// TIA Portal project "项目8" (V15.1)

(* hardware
DEVICE "GSD device_1"  GSD.Device.PN
   slot 0: "机架"  Rack  V1.0
   slot 0: "SINAMICS-G120SV-PN"  SINAMICS G120 CU250S-2 PN Vector V4.7  6SL3 246-0BA22-1FAx  V4.70
      slot 0: "SINAMICS G120 CU250S-2 PN Vector V4.7"  SINAMICS G120 CU250S-2 PN Vector V4.7
      slot 1: "DO 矢量_1"  DO VECTOR
         slot 0: "模块访问点"  Module Access Point
      slot 1: "PN-IO"  PN-IO
         slot 1: "端口1"  Port 1
         slot 2: "端口2"  Port 2
   slot 2: "标准报文1, PZD-2/2"  Standard telegram 1, PZD-2/2
DEVICE "S7-1200 station_1"  S7-1200 Station
   slot 0: "Rack_0"  S7-1200 Rack  Rack  V1.0
   slot 1: "PLC_1"  CPU 1214C DC/DC/DC  6ES7 214-1AG40-0XB0  V4.2
   slot 2: "DI 16/DQ 16x24VDC_1"  6ES7 223-1BL32-0XB0  V2.0
   slot 3: "AI 4x13BIT/AQ 2x14BIT_1"  6ES7 234-4HE32-0XB0  V2.0
DEVICE "HMI_1"  KTP700 Basic PN
   slot 0: "HMI_1"  KTP700 Basic PN  6AV2 123-2GB03-0AX0  15.1.0.0
   slot 1: "HMI_RT_1"  KTP700 Basic PN  6AV2 123-2GB03-0AX0  15.1.0.0
   slot 5: "HMI_1.IE_CP_1"  PROFINET Interface  15.0.1.0
      slot 1: "PROFINET Interface_1"  PROFINET Interface
         slot 1: "Port_1"  Port
*)

// ===== PLC "PLC_1"  CPU 1214C DC/DC/DC =====

VAR_GLOBAL   // PLC tag table "默认变量表"
   "G120输出速度" AT %MW0 : Word;
   "G120控制" AT %QW64 : Word;
   "Tag_5" AT %MW12 : Word;
   "G120速度" AT %QW66 : Word;
   "停止" AT %I0.1 : Bool;
   "正转" AT %I0.2 : Bool;
   "反转" AT %I0.3 : Bool;
   "轴_1_脉冲" AT %Q0.0 : Bool;
   "轴_1_方向" AT %Q0.1 : Bool;
   "开关4" AT %I0.4 : Bool;
   "步进电机启动" AT %Q1.0 : Bool;
   "速度" AT %MD10 : Real;
   "32位速度" AT %MD14 : DInt;
   "16位速度" AT %MW18 : UInt;
   "计算速度" AT %MD20 : Real;
   "sds" AT %MW24 : Int;
END_VAR

DATA_BLOCK "轴_1"   // DB1, Motion_DB
{ S7_Optimized_Access := 'TRUE' }
AUTHOR : SIMATIC
FAMILY : BasicMC
NAME : TO_PosAx
VERSION : 6.0
// stored: InstanceOfName TO_PositioningAxis
"TO_PositioningAxis"
BEGIN
   // Axis.LengthUnit.LastDistance = 1005
   // Axis.LengthUnitNormalized.Distance = 1005
   // Axis.DirectionOutputEnabledCU = TRUE
   // Axis.OnlinePtoModeCU = 16#0000_0002
   // Axis.SelectedChannel2EnumCU = %Q0.1
   // Axis.SelectedChannel1EnumCU = %Q0.0
   // Pulse.MinDeltaDeltaFrequencyCU = 0.004
   // Pulse.MaxDeltaDeltaFrequencyCU = 1.0E+10
   // Pulse.MinDeltaFrequencyCU = 0.005
   // Pulse.MaxDeltaFrequencyCU = 9.5E+9
   // Pulse.MinFrequencyCU = 1.0
   // Pulse.MaxFrequencyCU = 100000.0
   // Pulse.OutputSourceCU = 16#0000_0000
   // Axis.SelectPTO = 0
END_DATA_BLOCK

ORGANIZATION_BLOCK "Main"   // OB1, LAD, ProgramCycle
TITLE = "Main Program Sweep (Cycle)"
{ S7_Optimized_Access := 'TRUE' }
VERSION : 0.1
   VAR_INPUT
      Initial_Call : Bool;   // Initial call of this OB
      Remanence : Bool;   // =True, if remanent data are available
   END_VAR
BEGIN

REGION Network 1
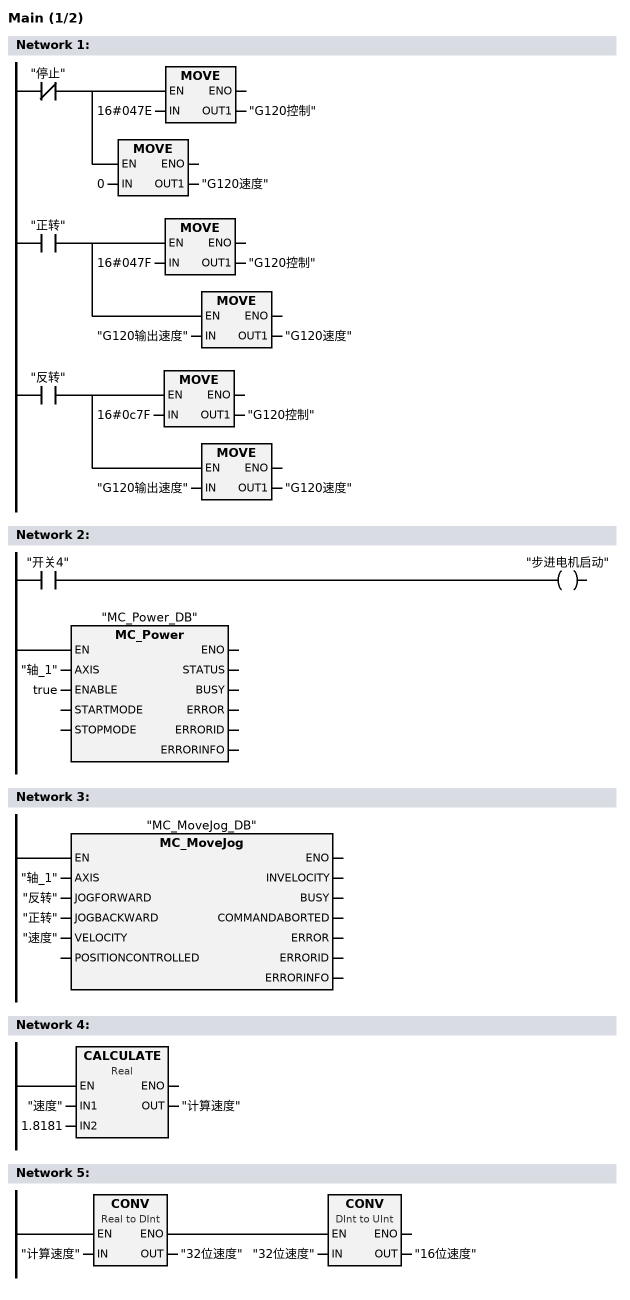
   RUNG wire#powerrail
      I_Contact( "停止" )
      wire#w1
      Move(in := 16#047E, out1 => "G120控制")
   END_RUNG
   RUNG wire#w1
      Move(in := 0, out1 => "G120速度")
   END_RUNG
   RUNG wire#powerrail
      Contact( "正转" )
      wire#w2
      Move(in := 16#047F, out1 => "G120控制")
   END_RUNG
   RUNG wire#w2
      Move(in := "G120输出速度", out1 => "G120速度")
   END_RUNG
   RUNG wire#powerrail
      Contact( "反转" )
      wire#w3
      Move(in := 16#0c7F, out1 => "G120控制")
   END_RUNG
   RUNG wire#w3
      Move(in := "G120输出速度", out1 => "G120速度")
   END_RUNG
   // the same network as SCL:
   IF NOT "停止" THEN
       "G120控制" := 16#047E;
       "G120速度" := 0;
   END_IF;
   IF "正转" THEN
       "G120控制" := 16#047F;
       "G120速度" := "G120输出速度";
   END_IF;
   IF "反转" THEN
       "G120控制" := 16#0c7F;
       "G120速度" := "G120输出速度";
   END_IF;
END_REGION

REGION Network 2
   "步进电机启动" := "开关4";
   "MC_Power_DB"(Axis := "轴_1", Enable := true);   // MC_Power
END_REGION

REGION Network 3
   "MC_MoveJog_DB"(Axis := "轴_1", JogForward := "反转", JogBackward := "正转", Velocity := "速度");   // MC_MoveJog
END_REGION

REGION Network 4
   RUNG wire#powerrail
      { S7_Templates := "SrcType := Real"; S7_Expression := "IN1*IN2" } Calculate(in1 := "速度", in2 := 1.8181, out => "计算速度")
   END_RUNG
   // the same network as SCL:
   "计算速度" := "速度"*1.8181;
END_REGION

REGION Network 5
   RUNG wire#powerrail
      { S7_Templates := "[SrcType := Real, DestType := DInt]" } Convert(in := "计算速度", out => "32位速度")
      { S7_Templates := "[SrcType := DInt, DestType := UInt]" } Convert(in := "32位速度", out => "16位速度")
   END_RUNG
   // the same network as SCL:
   "32位速度" := REAL_TO_DINT("计算速度");
   "16位速度" := DINT_TO_UINT("32位速度");
END_REGION

REGION Network 6
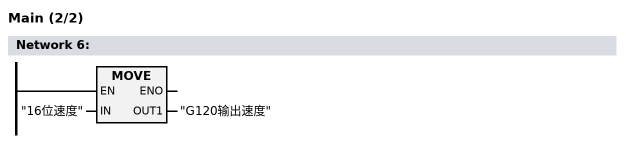
   RUNG wire#powerrail
      Move(in := "16位速度", out1 => "G120输出速度")
   END_RUNG
   // the same network as SCL:
   "G120输出速度" := "16位速度";
END_REGION
END_ORGANIZATION_BLOCK

ORGANIZATION_BLOCK "Startup"   // OB100, SCL, Startup
TITLE = "Complete Restart"
{ S7_Optimized_Access := 'TRUE' }
VERSION : 0.1
   VAR_INPUT
      LostRetentive : Bool;   // True if retentive data are lost
      LostRTC : Bool;   // True if date and time are lost
   END_VAR
BEGIN
   "速度" := 150;
END_ORGANIZATION_BLOCK

(* ===== HMI "HMI_RT_1" =====
system functions are stored by id; their names below are inferred from use
connection "HMI_连接_1": ETHERNET, SMART_S7_1200_OMS

HMI tags "默认变量表"
   "Tag_ScreenNumber" : UInt, internal
   "Tag_3" : Real = PLC 速度 AT %MD10, 1 s

Template "模板_1" 800x480
   Button "退出" at 714,429 size 71x50; TextOff '退出'; PictureOff "ExitRuntime_KTP700_Basic_PN_TR"; PictureOn "ExitRuntime_KTP700_Basic_PN_TR"
      on Release: StopRuntime(0)
   Button "Template_Button" at 614,429 size 71x50; TextOff 'Text'
   Button "Template_Button_1" at 514,429 size 71x50; TextOff 'Text'
   Button "Template_Button_2" at 414,429 size 71x50; TextOff 'Text'
   Button "Template_Button_3" at 314,429 size 71x50; TextOff 'Text'
   Button "Template_Button_4" at 214,429 size 71x50; TextOff 'Text'
   Button "Template_Button_5" at 114,429 size 71x50; TextOff 'Text'
   Button "起始画面" at 14,429 size 71x50; TextOff '起始画面'; PictureOff "NavigateHome_KTP700_Basic_PN_TR"; PictureOn "NavigateHome_KTP700_Basic_PN_TR"
      on Release: ActivateScreen("根画面", 0)
   SymbolicIOField "Symbolic_IO_Field_Screen" at 93,9 size 600x33; TextOff '0'; TextOn '1'; TextList "TextList_ScreenNames"
      ProcessValue <- "Tag_ScreenNumber"
      on Change: ActivateScreenByNumber("Tag_ScreenNumber", 0)
   DateTimeField "HmiScreenItemData" at 695,25 size 105x25
   DateTimeField "HmiScreenItemData_1" at 695,0 size 105x25
   GraphicView "Logo" at 0,0 size 91x51; Picture "HMI_1 的 Logo"

screen "根画面" 800x480, template "模板_1"
   on GenerateScreen: SetTag("Tag_ScreenNumber", 1)
   TextField "HmiScreenItemData" at 80,225 size 640x25; Text '欢迎进入 HMI_1 (KTP700 Basic+ PN)！'
   IOField "I/O 域_1" at 39,217 size 716x168; FormatPattern 999999999.999
      ProcessValue <- "Tag_3"
   TextField "文本域_1" at 295,94 size 199x101; Text '速度'
*)